(* IEC 61131-3 sources: plcassist-cli/packages/volt-lsp-iec/test-corpus/bakon-nano/Device/Plc Logic/Application/Library Manager/SysDir, 13 files *)

(* ---- DIRINFOFLAGS.gvl ---- *)
VAR_GLOBAL
	DF_FILE : DWORD := 16#0;
	DF_DIRECTORY : DWORD := 16#2;
END_VAR

(* ---- GVL.gvl ---- *)
VAR_GLOBAL
	SYSDIR_INVALID_HANDLE : RTS_IEC_HANDLE := RTS_INVALID_HANDLE;
END_VAR

(* ---- SYSDIRCLOSE.fun ---- *)
FUNCTION SYSDIRCLOSE : RTS_IEC_RESULT
VAR_INPUT
	HDIR : RTS_IEC_HANDLE;
END_VAR
END_FUNCTION

(* ---- SYSDIRCOPY.fun ---- *)
FUNCTION SYSDIRCOPY : RTS_IEC_RESULT
VAR_INPUT
	SZDESTDIR : REFERENCE TO STRING;
	SZSOURCEDIR : REFERENCE TO STRING;
	XRECURSIVE : BOOL;
	XOVERWRITE : BOOL;
END_VAR
END_FUNCTION

(* ---- SYSDIRCREATE.fun ---- *)
FUNCTION SYSDIRCREATE : RTS_IEC_RESULT
VAR_INPUT
	SZDIR : REFERENCE TO STRING;
END_VAR
END_FUNCTION

(* ---- SYSDIRCREATE2.fun ---- *)
FUNCTION SYSDIRCREATE2 : RTS_IEC_RESULT
VAR_INPUT
	SZDIR : REFERENCE TO STRING;
	XRECURSIVE : BOOL;
END_VAR
END_FUNCTION

(* ---- SYSDIRDELETE.fun ---- *)
FUNCTION SYSDIRDELETE : RTS_IEC_RESULT
VAR_INPUT
	SZDIR : REFERENCE TO STRING;
END_VAR
END_FUNCTION

(* ---- SYSDIRDELETE2.fun ---- *)
FUNCTION SYSDIRDELETE2 : RTS_IEC_RESULT
VAR_INPUT
	SZDIR : REFERENCE TO STRING;
	XRECURSIVE : BOOL;
	XKEEPDIR : BOOL;
END_VAR
END_FUNCTION

(* ---- SYSDIRGETCURRENT.fun ---- *)
FUNCTION SYSDIRGETCURRENT : RTS_IEC_RESULT
VAR_INPUT
	DIMAXDIRLEN : DINT;
END_VAR
VAR_IN_OUT
	SZDIR : STRING;
END_VAR
END_FUNCTION

(* ---- SYSDIROPEN.fun ---- *)
FUNCTION SYSDIROPEN : RTS_IEC_HANDLE
VAR_INPUT
	SZDIR : REFERENCE TO STRING;
	SZDIRENTRY : REFERENCE TO STRING;
	DIMAXDIRENTRY : DINT;
	PDIRINFO : POINTER TO DirInfo;
	PRESULT : POINTER TO RTS_IEC_RESULT;
END_VAR
END_FUNCTION

(* ---- SYSDIRREAD.fun ---- *)
FUNCTION SYSDIRREAD : RTS_IEC_RESULT
VAR_INPUT
	HDIR : RTS_IEC_HANDLE;
	DIMAXDIRENTRY : DINT;
	PDIRINFO : POINTER TO DirInfo;
END_VAR
VAR_IN_OUT
	SZDIRENTRY : STRING;
END_VAR
END_FUNCTION

(* ---- SYSDIRRENAME.fun ---- *)
FUNCTION SYSDIRRENAME : RTS_IEC_RESULT
VAR_INPUT
	SZOLDDIRNAME : REFERENCE TO STRING;
	SZNEWDIRNAME : REFERENCE TO STRING;
END_VAR
END_FUNCTION

(* ---- SYSDIRSETCURRENT.fun ---- *)
FUNCTION SYSDIRSETCURRENT : RTS_IEC_RESULT
VAR_INPUT
	SZDIR : REFERENCE TO STRING;
END_VAR
END_FUNCTION
